(* IEC 61131-3 sources: 2026_Projet_YGO_ExcavatriceDragage/CODE_BACKUP/CODE_20260907_ChantierWeekEnd_v0.6.43/J_SUPERVISION/_TYPES/1_TREUILS_BENNE, 26 files *)

(* ---- E_WinchTraceBlockReason.st ---- *)
(* =======================================================================
   E_WinchTraceBlockReason - Cause de blocage priorisee treuil (trace terrain)
   -----------------------------------------------------------------------
   Role : Ordre de priorite de la cause de blocage d'un treuil M1/M2,
      calcule en PRG_04_Treuils_Benne (#8bis) et publie via Data.TraceM1/M2.
      L'ordre de l'enum EST l'ordre de priorite (valeur croissante = priorite
      decroissante) : la cause la plus grave gagne (PowerCutOff > ... > NONE).
   Producteur unique : PRG_04_Treuils_Benne (#8bis).
   Consommateur : FB_TroubleshootingView (recopie -> GVL_Troubleshooting.TraceM1/2).
   Lecture seule - aucune action de conduite n'en depend.
   Doc metier : DOC/AF/AF_Partie-14_Fonction_Troubleshooting_v1.4.md
   ======================================================================= *)
{attribute 'qualified_only'}
TYPE E_WinchTraceBlockReason :
(
    NONE                    := 0,   // Aucun blocage - au moins un sens effectivement permis
    POWER_CUTOFF            := 1,   // Coupure puissance amont (instSafetyWinch.PowerCutOff) - priorite max
    AXIS_DISABLED           := 2,   // Axe neutralise (Mode=DISABLE ou InhibitMx -> Enable FALSE)
    SAFESTOP                := 3,   // SafeStop effectif (rampe rapide demandee)
    SAFETY_FAULT            := 4,   // Defaut safety latched (FB_Safety_Winch.Fault.Error)
    SAFETY_PERMIT_MISSING   := 5,   // Aucun sens ne delivre de permit safety (limite / mou de cable / homing)
    PROCESS_PERMIT_MISSING  := 6,   // Permit process absent (benne / fond Kobold / limite legale / extraction)
    COUPLING_BLOCKED        := 7,   // Couplage synchro anti-telescopage (l'autre axe bloque)
    WINCH_FAULT             := 8,   // Defaut treuil latched (FB_Winch.Fault.Error)
    FINAL_INTERLOCK_BLOCKED := 9    // Barriere finale en defaut (frein / redemarrage)
);
END_TYPE

(* ---- ST_BucketCfg.st ---- *)
(* ═══════════════════════════════════════════════════════════════
   ST_BucketCfg — Configuration de la benne (M2)
   ═══════════════════════════════════════════════════════════════ *)
TYPE ST_BucketCfg :
STRUCT
    Config              : ST_fbBucket_Config; (* Offsets Open/Close/Coherence *)
    CfgTimeoutDuration  : TIME := T#30s;    (* ⏱️ Temps max pour l'ouverture/fermeture *)
    Initialized         : BOOL := FALSE;   (* 🚦 flag restauration boot *)
END_STRUCT
END_TYPE

(* ---- ST_BucketCmd.st ---- *)
(* ═══════════════════════════════════════════════════════════════
   🎮 ST_BucketCmd — Commandes IHM pour la benne (M2)
   ═══════════════════════════════════════════════════════════════ *)
TYPE ST_BucketCmd :
STRUCT
    BtnOpen             : BOOL; (* 🪣 Bouton commande ouverture *)
    BtnClose            : BOOL; (* 🪣 Bouton commande fermeture *)
    BtnReset            : BOOL; (* 🔑 Acquittement défaut benne *)
    BtnConfirmOpenPos   : BOOL; (* Référencement benne position ouverte (mise en service) — confirmation pure, aucun mouvement *)
    BtnConfirmClosePos  : BOOL; (* Référencement benne position fermée (mise en service) — confirmation pure, aucun mouvement *)
    // Mode pilotage unitaire M2 "sécurisé" -- actif
    // uniquement en SelJoystickWinch=2 (unitaire M2). Si TRUE : borne le déplacement entre les
    // positions ouvert/fermé configurées (OffsetOpenM/OffsetCloseM relatif à M1, mêmes bornes que
    // FB_Bucket) ET plafonne la vitesse au palier 1, sans passer par instBucket (pas de mémorisation
    // CloseReq/OpenReq, jogging libre borné). Défaut FALSE : pilotage unitaire M2 sans limite dédiée.
    TglManualBucketLimits : BOOL := TRUE; // Défaut TRUE -- pilotage unitaire M2 borné + palier 1 par défaut
    // Assistance "vidage à la trémie" (MAINT_N1/N2) : arme l'ouverture auto de la benne quand
    // M3 est stable à la Trémie. Indépendant du verrou descente treuil (WinchDescentAuth_M3).
    TglEnableDumpAtTremie : BOOL := FALSE;
END_STRUCT
END_TYPE

(* ---- ST_BucketHMI.st ---- *)
(* ═══════════════════════════════════════════════════════════════
   ⚙️ ST_BucketHMI — Données d'échange IHM pour la benne (M2)
   ───────────────────────────────────────────────────────────────
   📄 Structuration en Cmd / State / Cfg / Bypass , homogène avec ST_WinchHMI.
   ═══════════════════════════════════════════════════════════════ *)
TYPE ST_BucketHMI :
STRUCT
    Cmd    : ST_BucketCmd;
    State  : ST_BucketHMIState;
    Cfg    : ST_BucketCfg;
    Bypass : ST_BypassBucket;
END_STRUCT
END_TYPE

(* ---- ST_BypassBucket.st ---- *)
(* ═══════════════════════════════════════════════════════════════
   ST_BypassBucket — Bypass de la surveillance benne (M2)
   🔒 Doctrine : actionnable UNIQUEMENT en MAINT_N2, RETAIN, jamais masque
      les autres défauts du même bloc.
   ═══════════════════════════════════════════════════════════════ *)
TYPE ST_BypassBucket :
STRUCT
    (* 🛡️ 1. Hiérarchie & Restauration *)
    Global      : BOOL; (* 🌐 Bypass Global : ignore toute surveillance du mécanisme benne *)
    // Flag restauration boot dédié (défaut FALSE non ambigu, contrairement à une valeur métier)
    Initialized : BOOL := FALSE; (* 🚦 TRUE = bypass restauré depuis GVL_BypassRetain ce boot *)
END_STRUCT
END_TYPE

(* ---- ST_BypassWinch.st ---- *)
(* ═══════════════════════════════════════════════════════════════
   ST_BypassWinch — Bypass maintenance dédiés à UN treuil (M1 ou M2)
   ───────────────────────────────────────────────────────────────
   🎨 Regroupe les bypass "dégradé assumé" propres à un axe (codeur,
      contacteurs) — chaque treuil a son propre matériel, donc son
      propre struct (imbriqué M1Winch.Bypass / M2Winch.Bypass).
   🔒 Doctrine : actionnable UNIQUEMENT en MAINT_N2, RETAIN, jamais masque
      les autres défauts du même bloc (voir REGISTRE_ACTIONS_Bypass_v1.0 (archive)).
   ⚠️ Les bypass de capteurs COMMUNS (SlackCable, TopPositionSensor — capteur
      physique unique partagé M1/M2) sont dans ST_CommunHMI.Bypass, PAS ici.
   ═══════════════════════════════════════════════════════════════ *)
TYPE ST_BypassWinch :
STRUCT
    (* 📡 1. Communication & Systèmes auxiliaires *)
    OperatorComm      : BOOL; (* 📡 Bypass communication esclave CANopen Joystick / heartbeat IHM *)
    EncoderFault      : BOOL; (* 🔌 Bypass diagnostic esclave EtherCAT COD (codeur absolu) *)
    ContactorFeedback : BOOL; (* 🔌 Bypass feedbacks contacteurs de puissance et frein *)
    PhaseRotation     : BOOL; (* ⚡ Bypass défaut rotation de phases (commun machine) *)
    BrakeThermal      : BOOL; (* 🌡️ Bypass surchauffe thermique frein (commun machine) *)
    MotorThermal      : BOOL; (* : 🌡️ Bypass surchauffe thermique moteur CE treuil (M1_ThermalOk_DI/M2_ThermalOk_DI) *)

    (* 🚧 2. Limites physiques et Positionnement *)
    TopLimitSwitch    : BOOL; (* 🚧 Bypass fin de course physique haute (capteur, bit5) *)
    TopLimitSoftware  : BOOL; (* : Bypass fin de course logiciel haut (position calculée CablePosM >= TopLimitM, symétrique CableLimitSwitch) *)
    CableLimitSwitch  : BOOL; (* 🚧 Bypass limite basse physique (longueur de câble max) *)
    LimitLegal        : BOOL; (* : Bypass limite légale de profondeur (GVL_IHM.Commun.LimitLegalReached) *)

    (* ⚙️ 3. Sécurité Mécanique (Méca A-E) *)
    MecaA             : BOOL; (* 🔄 Bypass Méca A : mouvement non commandé à l'arrêt *)
    MecaB             : BOOL; (* 🛑 Bypass Méca B : absence confirmation arrêt (frein/contacteurs) *)
    MecaC             : BOOL; (* 🏋️ Bypass Méca C : glissement de charge (benne M1) *)
    MecaD             : BOOL; (* 🚧 Bypass Méca D : arrivée butée haute anormale *)
    MecaE             : BOOL; (* 🔄 Bypass Méca E : désynchronisation critique *)

    (* 🛡️ 4. Hiérarchie & Restauration *)
    Safety            : BOOL; (* 🛡️ Bypass groupé : tous les bits qui provoquent un PowerCutOff *)
    Process           : BOOL; (* ⚙️ Bypass groupé : tous les bits qui provoquent un SafeStop *)
    Global            : BOOL; (* 🌐 Bypass Global : ignore toutes les sécurités de cet axe *)
    // Flag restauration boot dédié (défaut FALSE non ambigu, contrairement à une valeur métier)
    Initialized       : BOOL := FALSE; (* 🚦 TRUE = bypass restauré depuis GVL_BypassRetain ce boot *)
END_STRUCT
END_TYPE

(* ---- ST_Chain_Winch_Control.st ---- *)
TYPE ST_Chain_Winch_Control :
STRUCT
    Idx401_MotionAllowed         : BOOL; // 1 = Prêt / Mouvement Autorisé | 0 = Bloqué
    Idx402_SpeedStepCalculated   : INT;  // Palier Vitesse Calculé (0, 1, 2, 3, 4)
    Idx403_SpeedRamp_Pct         : REAL; // [%] Consigne Vitesse après Rampe
    Idx404_BrakeReleaseAuthorized: BOOL; // 1 = Ordre Ouverture Frein | 0 = Ordre Serrage
    Idx405_FinalInterlockState   : E_WinchFinalInterlockState; // 🛡️ État frontière
    Idx406_FinalInterlockReason  : E_WinchFinalInterlockReason; // 🛡️ Cause mémorisée
    Idx407_FinalAuthorizedStep   : INT;  // 🪜 Palier réellement autorisé
    Idx408_BrakeCommandOpenConfirmed : BOOL; // 🔌 Contacteur/bobine, pas frein mécanique
    Idx409_BrakeTimeoutElapsed   : TIME; // ⏱️ Watchdog 500ms écoulé
    Idx410_RestartDelayElapsed   : TIME; // ⏱️ Verrou 900ms écoulé
    Idx411_StepDelayElapsed      : TIME; // ⏱️ Délai palier 1s250 écoulé
    Idx412_InTopSlowdownZone     : BOOL; // 🐢 Palier plafonné à 1, approche limite haute
    Idx413_InBottomSlowdownZone  : BOOL; // 🐢 Palier plafonné à 1, approche limite basse (câble ou légale)
    Idx414_BottomLimitActiveM    : REAL; // : Limite basse active (m) — câble physique OU légale, la plus restrictive
    (* 🔎 Diagnostic anti-redémarrage — "commande active mais rien ne tourne" *)
    Idx415_MotorRequest          : BOOL; // 1 = demande moteur active (palier>0 ET un seul sens) | 0 = pas de demande vue par la barrière
    Idx416_RestartRequired       : BOOL; // 1 = purge anti-redémarrage armée, AuthorizedStep force a 0 tant que non purgee
    Idx417_RestartInhibit        : BOOL; // 1 = verrou latché (frein non confirmé), exige Reset conscient — distinct de Idx416
    Idx418_NeutralRequestSeen    : BOOL; // 1 = passage au neutre observé pendant un RestartInhibit (réarmement en cours)
END_STRUCT
END_TYPE

(* ---- ST_Chain_Winch_Demandes.st ---- *)
TYPE ST_Chain_Winch_Demandes :
STRUCT
    Idx201_JoyRawPhysical_ANA    : INT;  // [pts] Bruts convertisseur (-2048 à +2048)
    Idx202_JoyScaledPhysical_Pct : REAL; // [%] Consigne Joystick (-100% à +100%)
    Idx203_HmiManualCmd_BtnAscent : BOOL; // 1 = Appui Bouton Ascending IHM | 0 = Relâché
    Idx204_HmiManualCmd_BtnDescent : BOOL; // 1 = Appui Bouton Descending IHM | 0 = Relâché
    Idx205_CycleAutoCmd_Pct      : REAL; // [%] Consigne auto envoyée par le Cycle
    Idx206_ModeActive            : E_Mode;// Mode courant (MANU_N1, AUTO_N1, MAINT_N2...)
    Idx207_BypassOperatorComm    : BOOL; // 0 = Comm Normale OK | 1 = Bypass Réseau Actif ⚠️
    Idx208_ArbitratedSpeed_Pct   : REAL; // [%] Consigne finale retenue après arbitrage
    Idx209_ArbitratedDirection   : INT;  // +1 = Ascending | 0 = Neutre | -1 = Descending
    Idx210_CoupledUserRequestDirection : INT; // +1 = Ascending | 0 = Neutre | -1 = Descending
    Idx211_CoupledUserRequestActive    : BOOL; // 1 = demande utilisateur couplée active
END_STRUCT
END_TYPE

(* ---- ST_Chain_Winch_Inputs.st ---- *)
TYPE ST_Chain_Winch_Inputs :
STRUCT
    Idx101_EncoderRawPos         : DINT; // [Valeur brutes pts] Codeur connecté
    Idx102_CablePos_M            : REAL; // [mètres] Position calculée du câble
    Idx103_ContactorsReleased_DI : BOOL; // 1 = OK (Tous contacteurs retombés à l'arrêt) | 0 = Contacteur collé
    Idx104_BrakeApplied          : BOOL; // TRUE = frein SERRÉ (NOT BrakeFeedback — IHM garde le sens serré)
    Idx105_ThermalOk_DI          : BOOL; // 1 = Température OK (Sain) | 0 = Surchauffe Moteur M1
END_STRUCT
END_TYPE

(* ---- ST_Chain_Winch_Outputs.st ---- *)
TYPE ST_Chain_Winch_Outputs :
STRUCT
    Idx501_CmdRelayAscent_DQ   : BOOL; // 1 = Relais Ascending ON | 0 = OFF
    Idx502_CmdRelayDescent_DQ  : BOOL; // 1 = Relais Descending ON | 0 = OFF
    Idx503_CmdSpeedContactor1_DQ : BOOL; // 1 = Contacteur Vitesse 1 ON | 0 = OFF
    Idx504_CmdSpeedContactor4_DQ : BOOL; // 1 = Contacteur Vitesse 4 ON (Plein Gaz) | 0 = OFF
    Idx505_CmdBrakeRelease_RQ    : BOOL; // 1 = Bobine Frein Alimentée (Ouvert) | 0 = Non Alimentée (Serré)
END_STRUCT
END_TYPE

(* ---- ST_Chain_Winch_Safety.st ---- *)
TYPE ST_Chain_Winch_Safety :
STRUCT
    Idx301_EmergencyChainClosed  : BOOL; // 1 = Boucle Urgence OK (Armé) | 0 = Arrêt d'Urgence Appuyé
    Idx302_SafeStopActive        : BOOL; // 0 = Sain (Autorisé) | 1 = Arrêt Rapide Métier Actif
    Idx303_PowerCutOffActive     : BOOL; // 0 = Puissance OK | 1 = Coupure Puissance Sécurité
    Idx304_TopSensorPhysical_DI  : BOOL; // 1 = Capteur Haut Libre (Sain) | 0 = Butée Haute Atteinte
    Idx305_TopSensorBypassActive : BOOL; // 0 = Capteur Actif | 1 = Capteur Haut Shunté IHM ⚠️
    Idx306_AscentPermitEffective  : BOOL; // 1 = Ascending Autorisée | 0 = ASCENDING BLOQUÉE
    Idx307_SlackCablePhysical_DI : BOOL; // 1 = Câble Tendu (Sain) | 0 = Mou de Câble Détecté
    Idx308_SlackCableBypassActive: BOOL; // 0 = Capteur Actif | 1 = Mou de Câble Shunté IHM ⚠️
    Idx309_DescendPermitEffective: BOOL; // 1 = Descending Autorisée | 0 = DESCENDING BLOQUÉE
    (* Défauts safety déchiffrés (bits ErrorId) — visibles individuellement à l'IHM *)
    Idx310_ErrorOperatorComm : BOOL; // bit0 Perte communication opérateur (joystick CAN / heartbeat IHM)
    Idx311_ErrorEncoder      : BOOL; // bit1 Perte codeur de ce treuil
    Idx312_ErrorPhaseRotation: BOOL; // bit4 Mauvaise rotation de phases
    Idx313_ErrorMecaA        : BOOL; // bit7 Mouvement non commandé / roue libre
    Idx314_ErrorMecaB        : BOOL; // bit8 Absence confirmation arrêt sans commande
    Idx315_ErrorMecaC        : BOOL; // bit9 Glissement M1 pendant cycle benne
    Idx316_ErrorMecaD        : BOOL; // bit11 Non-arrêt sur capteur haut
    Idx317_ErrorMecaE        : BOOL; // bit12/13 Écart synchro critique M1/M2
    Idx318_ErrorBrakeThermal : BOOL; // bit10 Surchauffe thermique frein commun
    Idx319_ErrorOppositeDir  : BOOL; // bit14 Sens réel opposé au sens commandé
    Idx320_ErrorNoMovement   : BOOL; // bit15 Absence de mouvement malgré commande
    (* ⛔ Bloc "Pourquoi la montée ne s'arrête pas à la limite haute ?" — diagnostic ordonné
       (lecture maintenance) : config + position → butée atteinte → bypass actifs. *)
    Idx321_CfgTopLimitM               : REAL;  // 📐 Limite haute effective active (m) = CfgCableLimitAscent_M
    Idx322_CablePosM                  : REAL;  // 📐 Position câble courante (m)
    Idx323_TopLimitReached            : BOOL;  // 1 = position >= limite haute (hors homing) | 0 = en dessous
    Idx324_AscentBlockedByTopLimit    : BOOL;  // 1 = montée réellement coupée par la butée logicielle (AscentPermit=0) | 0 = limitée non bloquante (bypass ?)
    Idx325_BypassTopLimitSoftware     : BOOL;  // ⚠️ 1 = butée logicielle shunétee IHM (individuel)
    Idx326_BypassTopLimitSoftCommun   : BOOL;  // ⚠️ 1 = butée logicielle shunétee (commun)
    Idx327_BypassTopLimitSwitch       : BOOL;  // ⚠️ 1 = capteur fin de course haut shuné IHM (individuel)
    Idx328_BypassTopLimitSwitchCommun : BOOL;  // ⚠️ 1 = capteur fin de course haut shuné (commun)
    Idx329_BypassGlobal               : BOOL;  // ⚠️ 1 = bypass global treuil (individuel)
    Idx330_BypassGlobalCommun         : BOOL;  // ⚠️ 1 = bypass global (commun)
END_STRUCT
END_TYPE

(* ---- ST_ChainBucket.st ---- *)
TYPE ST_ChainBucket :
STRUCT
    Idx101_BucketIsOpen          : BOOL; // 1 = Benne Mécaniquement Ouvert | 0 = Non Confirmé
    Idx102_BucketIsClosed        : BOOL; // 1 = Benne Mécaniquement Fermé | 0 = Non Confirmé
    Idx103_OffsetPos_M           : REAL; // [mètres] Écart d'Ouverture Câble M1/M2
    Idx104_AutoSeqActive         : BOOL; // : 1 = Séquencement auto (ouverture/fermeture armée par mouvement couplé) en cours
    Idx105_StateIncoherent       : BOOL; // : 1 = État ouvert/fermé INCONNU (ni IsOpen ni IsClosed fiable) -- cause fréquente de blocage
    Idx106_FBState               : E_State; // : État machine FB_Bucket (READY/BUSY/DONE/DISABLED)
    Idx107_LastPosM2Open_M       : REAL; // : Dernière position M2 mémorisée "ouvert"
    Idx108_LastPosM2Close_M      : REAL; // : Dernière position M2 mémorisée "fermé"
    Idx109_BucketTooOpen         : BOOL; // ⚠️ Dépassement ouverture : Delta < OffsetOpen - Tolerance (Enrouler M2)
    Idx110_BucketTooClosed       : BOOL; // ⚠️ Dépassement fermeture : Delta > OffsetClose + Tolerance (Dérouler M2)
    Idx111_BucketIsIntermediate  : BOOL; // ↔️ Position intermédiaire (entrebâillée entre ouvert et fermé)
    Idx112_DeltaPosition_M       : REAL; // 📏 Écart réel signé M2 - M1 (mètres) en direct

    Idx113_MachineHomed : BOOL; // Reference M1/M2/benne qualifiee
    Idx114_MachineHomingStep         : INT;  // Etape guidee reference machine
    Idx115_MachineHomingFailed       : BOOL; // Transaction reference abandonnee
    Idx116_M1ReferenceMissing    : BOOL; // M1 non reference ou mesure douteuse
    Idx117_M2ReferenceMissing    : BOOL; // M2 non reference ou mesure douteuse
    Idx118_BucketOffsetUnknown   : BOOL; // Offset benne non confirme
    Idx119_ReferenceTransaction  : BOOL; // Homing conjoint en cours
    Idx120_MachineHomingLossSafeStop : BOOL; // Perte reference pendant mouvement

    Idx201_HmiCmd_BtnOpen        : BOOL; // 1 = Demande Ouverture IHM | 0 = Relâché
    Idx202_HmiCmd_BtnClose       : BOOL; // 1 = Demande Fermeture IHM | 0 = Relâché
    Idx203_CycleCmd_Open         : BOOL; // 1 = Demande Ouverture par le Cycle Auto
    Idx204_CoupledDiveOpenArmed   : BOOL; // : 1 = Ouverture auto armée (descente couplée demandée, benne pas ouverte)
    Idx205_CoupledAscentCloseArmed: BOOL; // : 1 = Fermeture auto armée (montée couplée demandée, benne pas fermée)
    Idx206_CloseReqActive        : BOOL; // : 1 = Fermeture mémorisée/en cours (instBucket.CloseReq -- reste à 1 si recul partiel non terminé)
    Idx207_OpenReqActive         : BOOL; // : 1 = Ouverture mémorisée/en cours (instBucket.OpenReq -- idem)
    Idx208_MotionBlockedByBucket : BOOL; // : 1 = Mouvement couplé BLOQUÉ (auto-séquencement armé mais benne pas Busy -- vérifier Idx306_ErrorIdRaw)

    Idx301_EmergencyChainClosed  : BOOL; // 1 = Boucle Urgence OK | 0 = AU Appuyé
    Idx302_BucketFaultActive     : BOOL; // 0 = Sain | 1 = Défaut Mouvement Benne
    Idx303_KoboldAutoStopEnabled       : BOOL; // 1 = Toggle IHM arrêt auto descente actif
    Idx304_KoboldImmersionConfirmed    : BOOL; // : 1 = Immersion confirmée (front Kobold dans la fenêtre)
    Idx305_KoboldBottomTouchLatched    : BOOL; // : 1 = Fond détecté, descente bloquée (ProcessPermitM1/M2_Descend)
    Idx306_ErrorIdRaw             : WORD; // : bitfield brut FB_Bucket (bit0 configuration, bit1 écart M2/M1, bit2 timeout, bit3 glissement M1, bit4 codeurs non référencés)
    Idx307_EffectivePermit_Open    : BOOL; // 1 = ouverture benne physiquement autorisée
    Idx308_EffectivePermit_Close   : BOOL; // 1 = fermeture benne physiquement autorisée

    Idx401_BucketBusy            : BOOL; // 1 = Mouvement Mâchoires en cours | 0 = Repos
    Idx402_BucketDone            : BOOL; // 1 = Position Cible Atteinte | 0 = En cours
    Idx403_ExtractionControlActive : BOOL; // : 1 = Phase vitesse contrôlée montée en cours

    Idx501_M2_CmdRev_DQ          : BOOL; // 1 = Relais Action Benne M2 ON
END_STRUCT
END_TYPE

(* ---- ST_ChainWinch.st ---- *)
TYPE ST_ChainWinch :
STRUCT
    Inputs_100    : ST_Chain_Winch_Inputs;
    Demandes_200  : ST_Chain_Winch_Demandes;
    Safety_300    : ST_Chain_Winch_Safety;
    Control_400   : ST_Chain_Winch_Control;
    Outputs_500   : ST_Chain_Winch_Outputs;
END_STRUCT
END_TYPE

(* ---- ST_ChainWinchSync.st ---- *)
TYPE ST_ChainWinchSync :
STRUCT
    Idx101_M1_CablePos_M         : REAL; // [mètres] Position Câble M1 Retenue
    Idx102_M2_CablePos_M         : REAL; // [mètres] Position Câble M2 Benne
    Idx103_SyncDelta_M           : REAL; // [mètres] Écart Relatif M1 - M2

    Idx201_JoyYRaw_Pct           : REAL; // [%] Consigne Joystick Axe Y (-100% à +100%)
    Idx202_SyncEnabled_IHM       : BOOL; // 1 = Couplage Synchro Actif (Nominal) | 0 = Découplé ⚠️
    Idx203_ArbitratedSpeed_Pct   : REAL; // [%] Consigne Vitesse Synchro Arbitrée

    Idx301_EmergencyChainClosed  : BOOL; // 1 = Boucle Urgence OK | 0 = Arrêt Urgence
    Idx302_SyncFaultActive       : BOOL; // 0 = Synchro OK | 1 = Écart Synchro Bloquant
    Idx303_M1_AscentPermit       : BOOL; // 1 = Ascending M1 Autorisée | 0 = Bloquée (Fdc/Safety)
    Idx304_M2_AscentPermit       : BOOL; // 1 = Ascending M2 Autorisée | 0 = Bloquée (Fdc/Safety)

    Idx401_SyncMotionAllowed     : BOOL; // 1 = Mouvement Synchro Autorisé | 0 = Bloqué
    Idx402_M1_SetpointSpeed_Pct  : REAL; // [%] Consigne Vitesse Calculée M1
    Idx403_M2_SetpointSpeed_Pct  : REAL; // [%] Consigne Vitesse Calculée M2

    Idx501_M1_CmdRelayFwd_DQ     : BOOL; // 1 = Ascending M1 ON | 0 = OFF
    Idx502_M2_CmdRelayFwd_DQ     : BOOL; // 1 = Ascending M2 ON | 0 = OFF
END_STRUCT
END_TYPE

(* ---- ST_HwWinch.st ---- *)
(* ═══════════════════════════════════════════════════════════════
   🏗️ ST_HwWinch — Image matérielle brute des entrées Treuils M1 / M2
   ───────────────────────────────────────────────────────────────
   🎨 Regroupe les signaux physiques d'entrée bruts des treuils M1 et M2.
   ═══════════════════════════════════════════════════════════════ *)
TYPE ST_HwWinch :
STRUCT
    M1_ContactorsReleased_DI : BOOL; (* Retours contacteurs M1 retombés *)
    M1_ThermalOk_DI          : BOOL; (* Thermique moteur M1 OK *)
    M1_BrakeIsOpen_DI        : BOOL; (* Retour frein M1 (1 = ouvert) *)

    M2_ContactorsReleased_DI : BOOL; (* Retours contacteurs M2 retombés *)
    M2_ThermalOk_DI          : BOOL; (* Thermique moteur M2 OK *)
    M2_BrakeIsOpen_DI        : BOOL; (* Retour frein M2 (1 = ouvert) *)

    M1M2_TopPositionFree_DI  : BOOL; (* Capteur position haute commun M1/M2 libre *)
    M2_TensionedCable_DI     : BOOL; (* Capteur mou de câble M2 (câble tendu) *)

    COD1_PosValue            : UDINT;        (* Valeur brute position codeur COD1 (M1) *)
    COD1_SpdValue            : DINT;         (* Valeur brute vitesse codeur COD1 (0x6031:01 en 0.1 RPM) *)
    COD1_Alarms              : UINT;         (* Alarmes brutes COD1 *)
    COD1_Warnings            : UINT;         (* Avertissements bruts COD1 *)
    COD1_DeviceState         : DEVICE_STATE; (* État device COD1 (GetDeviceState) *)

    COD2_PosValue            : UDINT;        (* Valeur brute position codeur COD2 (M2) *)
    COD2_SpdValue            : DINT;         (* Valeur brute vitesse codeur COD2 (0x6031:01 en 0.1 RPM) *)
    COD2_Alarms              : UINT;         (* Alarmes brutes COD2 *)
    COD2_Warnings            : UINT;         (* Avertissements bruts COD2 *)
    COD2_DeviceState         : DEVICE_STATE; (* État device COD2 (GetDeviceState) *)
END_STRUCT
END_TYPE

(* ---- ST_OutputsInterPrg.st ---- *)
(* ═══════════════════════════════════════════════════════════════
   📤 ST_OutputsInterPrg — Bus d'échange inter-PRG produit par PRG_06_Outputs
   ───────────────────────────────────────────────────────────────
   🎯 Rôle : Encapsuler les ordres actionneurs finaux (M1/M2/M3, AU) produits
      par PRG_06_Outputs et rebouclés par FB_SimBench (instancié dans
      PRG_02_Acquisition) pour le banc de simulation intégré.
   📤 Producteur unique : PRG_06_Outputs (VAR_OUTPUT Data : ST_OutputsInterPrg).
   📄 Doc : DOC/AF/AF_Partie-06_Acquisition_Qualification_IO_v2.4.md §5
   🔌 Architecture : Bus de données typé — encapsulation des échanges inter-PRG.
   ═══════════════════════════════════════════════════════════════ *)

TYPE ST_OutputsInterPrg :
STRUCT
    // === 🪝 Ordres actionneurs finaux treuil M1 ===
    M1RelayFwd            : BOOL; // 🛗 Ordre contacteur montee treuil M1
    M1RelayRev            : BOOL; // 🛗 Ordre contacteur descente treuil M1
    M1SpeedContactor1     : BOOL; // 🔌 Ordre contacteur palier 1 treuil M1
    M1SpeedContactor2     : BOOL; // 🔌 Ordre contacteur palier 2 treuil M1
    M1SpeedContactor3     : BOOL; // 🔌 Ordre contacteur palier 3 treuil M1
    M1SpeedContactor4     : BOOL; // 🔌 Ordre contacteur palier 4 treuil M1
    M1BrakeCmd            : BOOL; // 🔓 Ordre desserrage frein M1 (1=Desserrer)

    // === 🪝 Ordres actionneurs finaux treuil M2 ===
    M2RelayFwd            : BOOL; // 🛗 Ordre contacteur montee/fermeture treuil M2
    M2RelayRev            : BOOL; // 🛗 Ordre contacteur descente/ouverture treuil M2
    M2SpeedContactor1     : BOOL; // 🔌 Ordre contacteur palier 1 treuil M2
    M2SpeedContactor2     : BOOL; // 🔌 Ordre contacteur palier 2 treuil M2
    M2SpeedContactor3     : BOOL; // 🔌 Ordre contacteur palier 3 treuil M2
    M2SpeedContactor4     : BOOL; // 🔌 Ordre contacteur palier 4 treuil M2
    M2BrakeCmd            : BOOL; // 🔓 Ordre desserrage frein M2 (1=Desserrer)

    // === 🔀 Concordance contacteurs M1/M2 (instance FB_SyncContactor sur vecteurs finaux) ===
    ContactorMismatch          : BOOL;                  // Niveau 1 confirmé (debounce 500 ms) → SafeStop des 2 treuils (PRG_04, scan N-1)
    ContactorMismatchEscalated : BOOL;                  // Niveau 2 persistant → escalade PowerCutOff via latch MecaE (PRG_04)
    SyncContactorDiag          : ST_SyncContactorDiag;  // Détail : quel contacteur diverge + niveau atteint (IHM / troubleshooting)

    // === ↔️ Ordre actionneur final translation M3 ===
    TranslationBrakeCmd   : BOOL; // 🔓 Demande frein M3 arbitree

    // === 🚨 Chaîne réarmement puissance AU ===
    PowerKeepAliveACmd    : BOOL; // 🔒 Maintien puissance voie A (1=Maintenu)
    PowerKeepAliveBCmd    : BOOL; // 🔒 Maintien puissance voie B (1=Maintenu)
    EmergencyArmingCmd    : BOOL; // 🎯 Impulsion rearmement puissance AU
    TestCutActive         : BOOL; // 🧪 Test de redondance AU en cours (canal A ou B coupe) — consommé par FB_SimBench
    PowerCutOffRequest    : BOOL; // 🛑 Requête coupure métier (arrêt d'urgence) — consommé par FB_SimBench
END_STRUCT
END_TYPE

(* ---- ST_SafetyWinch.st ---- *)
(* ═══════════════════════════════════════════════════════════════
   🛡️ ST_SafetyWinch — Diagnostics de sécurité pour un treuil
   ───────────────────────────────────────────────────────────────
   🎨 Destiné à l'affichage des défauts de sécurité d'un treuil.
   ═══════════════════════════════════════════════════════════════ *)
TYPE ST_SafetyWinch :
STRUCT
    Error             : BOOL;    (* 🛡️ Bloc sécurité (Safety) en défaut *)
    ErrorId           : WORD;    (* ❌ Code bitfield du défaut de sécurité (vue LIVE) *)
    LatchedId         : WORD;    (* 🕘 Vue LATCHÉE : ErrorId figé au défaut, effacé au Reset (marqueur [HISTO]) *)
    SafeStop          : BOOL;    (* 🟧 Arrêt rapide activé par la sécurité *)
    DescendPermit     : BOOL;    (* 🟢 Descending autorisée (TRUE = OK | FALSE = mou de câble / limite basse) *)
    AscentPermit      : BOOL;    (* 🟢 Ascending autorisée (TRUE = OK | FALSE = fin de course haut) *)
    SlackCable        : BOOL;    (* ⚠️ Mou de câble physiquement détecté *)
    ThermalFault      : BOOL;    (* 🔥 Surchauffe thermique moteur *)
    EncoderFault      : BOOL;    (* 🔌 Perte de liaison ou incohérence codeur *)
    BypassActive      : BOOL;    (* Bypass codeur effectivement accepté, uniquement MAINT_N2 *)
    CableLimitDescent : BOOL;    (* ⚠️ Longueur max de câble atteinte (limite basse physique) *)
    CableLimitAscent  : BOOL;    (* ⚠️ Limite haute d'exploitation normale atteinte *)
    MecaADrift_M      : REAL;    (* 📐 Dérive mesurée Méca A (m) *)
    MecaCDrift_M      : REAL;    (* 📐 Dérive mesurée Méca C (m) *)
    MecaBElapsedTime  : TIME;    (* ⏳ Temps écoulé confirmation contacteurs/frein *)
    PowerCutOff       : BOOL;    (* 🧨 Coupure puissance amont activée *)
    BlockedBySafety   : BOOL;    (* 🚫 Synthèse globale : actionneur bloqué par la sécurité (PowerCutOff OU SafeStop/Error) *)
    PowerCutOffSafety : BOOL;    (* 🧨 Synthèse sécurités critiques entraînant une coupure puissance *)
    SafeStopSafety    : BOOL;    (* 🛡️ Synthèse défauts entraînant un SafeStop / Rampe rapide *)
    (* 🔍 Décomposition individuelle des défauts de sécurité (bits ErrorId) *)
    ErrorOperatorComm : BOOL;    (* 🎮 Perte communication opérateur : joystick CAN ou heartbeat IHM (bit0) *)
    ErrorEncoder      : BOOL;    (* 🔌 Perte de liaison ou incohérence codeur (bit1) *)
    ErrorPhaseRotation: BOOL;    (* ⚡ Mauvaise rotation de phases électriques (bit4) *)
    ErrorBrakeThermal : BOOL;    (* 🌡️ Surchauffe thermique frein commun M1/M2/M3 (bit10) *)
    ErrorMecaA        : BOOL;    (* 🔄 Mouvement non commandé / roue libre (Méca A - bit7) *)
    ErrorMecaB        : BOOL;    (* 🛑 Absence confirmation arrêt sans commande (Méca B - bit8) *)
    ErrorMecaC        : BOOL;    (* 🏋️ Glissement M1 pendant cycle benne (Méca C - bit9) *)
    ErrorMecaD        : BOOL;    (* 🚧 Non-arrêt sur capteur haut (Méca D - bit11) *)
    ErrorMecaE        : BOOL;    (* 🔄 Écart de synchronisation critique M1/M2 (Méca E - bit12/13) *)
    ErrorOppositeDir  : BOOL;    (* 🧭 Sens réel opposé au sens commandé (bit14) *)
    ErrorNoMovement   : BOOL;    (* ⏱️ Absence de mouvement malgré commande (bit15) *)
    ErrorOverspeed    : BOOL;    (* ⚡ Survitesse treuil mesurée au-delà du palier 5 (latchée, acquittée au Reset) *)
END_STRUCT
END_TYPE

(* ---- ST_TraceWinch.st ---- *)
(* =======================================================================
   ST_TraceWinch - Trace de blocage terrain d'un treuil M1/M2
   -----------------------------------------------------------------------
   Role : Publier au technicien une vue consolidee "pourquoi l'axe ne bouge
   pas" : permis effectifs par sens, source du SafeStop/coupure, cause de
   blocage priorisee et horodatee.
   Producteur unique : PRG_04_Treuils_Benne (#8bis) - 1 instance par axe
       (TraceM1 / TraceM2 au sein de ST_WinchInterPrg).
   Consommateur : FB_TroubleshootingView (pure recopie -> GVL_Troubleshooting).
   Lecture seule - aucun calcul de commande n'en depend.
   BlockReasonTimestamp : ms depuis demarrage PLC (TIME()), latched au dernier
       changement de BlockReason (1 scan, memoire).
   Doc metier : DOC/AF/AF_Partie-14_Fonction_Troubleshooting_v1.4.md
   ======================================================================= *)
TYPE ST_TraceWinch :
STRUCT
    // Permis effectifs par sens (reflet exact des permis appliques au mouvement)
    DescendPermitEffective  : BOOL;   // Descente effectivement permise (EffectivePermit*_Descend)
    AscentPermitEffective   : BOOL;   // Montee effectivement permise (EffectivePermit*_Ascent)
    AscentPermitApplied      : BOOL;   // Permis effectivement transmis a la barriere finale
    DescendPermitApplied     : BOOL;   // Permis effectivement transmis a la barriere finale
    FinalPermitBlocked       : BOOL;   // Demande presente mais refusee par le permis final

    // Source de SafeStop / coupure - pour distinguer l'origine du blocage
    SafeStopActive          : BOOL;   // SafeStop effectif applique (SafeStop*_Active)
    SafeStopSourceSafety    : BOOL;   // SafeStop issu de FB_Safety_Winch (defaut safety)
    SafeStopSourceInput     : BOOL;   // SafeStop issu du module d'entree / homing / slip benne
    SafeStopSourceSync      : BOOL;   // SafeStop issu de la synchro M1/M2 (couplage anti-telescopage)
    PowerCutOffActive       : BOOL;   // Coupure puissance amont active (instSafetyWinch.PowerCutOff)
    Inhibited               : BOOL;   // Axe neutralise (Mode=DISABLE ou InhibitMx)

    // Barriere finale (fin de course mecanique / frein / redemarrage)
    FinalInterlockError     : BOOL;   // Defaut barriere finale (frein / redemarrage)
    FinalInterlockReason    : E_WinchFinalInterlockReason; // Cause barriere finale memorisee

    // Cause de blocage priorisee + horodatage
    BlockReason             : E_WinchTraceBlockReason; // Cause de blocage prioritaire
    BlockReasonTimestamp    : UDINT;  // ms depuis demarrage PLC (TIME()) - dernier changement de BlockReason
    StepNumber              : INT;    // Palier de vitesse actif (WinchState.StepNumber)
END_STRUCT
END_TYPE

(* ---- ST_WinchBenneHMI.st ---- *)
(* ═══════════════════════════════════════════════════════════════
   ⚙️ ST_WinchBenneHMI — Données d'échange IHM pour le treuil Benne (M2 uniquement)
   ───────────────────────────────────────────────────────────────
   🎨 Composition dupliquée de ST_WinchHMI (Cmd/State/Cfg/Safety/Bypass) + Bucket.
   📄 IEC 61131-3 n'offre pas d'héritage de struct : cette duplication de la liste
      de champs est assumée pour garder M1TreuilRetenue (ST_WinchHMI, sans Bucket)
      strictement distinct de M2TreuilBenne (ce type, avec Bucket) — décision
      DOC/CHECKLISTS/TASK_CONTEXT/TASK_CONTEXT_LOT_TROUBLESHOOTING_VIEW_ET_WINCHHMI.yaml AC5.
   ═══════════════════════════════════════════════════════════════ *)
TYPE ST_WinchBenneHMI :
STRUCT
    (* 🎮 Commandes opérateur *)
    Cmd                     : ST_WinchCmd;

    (* 🚦 États, retours et mesures *)
    State                   : ST_WinchState;

    (* Configurations et limites *)
    Cfg                     : ST_WinchCfg;

    (* 🛡️ Sécurité (FB_Safety_Winch) *)
    Safety                  : ST_SafetyWinch;

    (* Bypass maintenance *)
    Bypass                  : ST_BypassWinch;

    (* 🪣 Benne — pertinent uniquement pour M2 (M2TreuilBenne.Bucket) *)
    Bucket                  : ST_BucketHMI;
END_STRUCT
END_TYPE

(* ---- ST_WinchCfg.st ---- *)
(* ═══════════════════════════════════════════════════════════════
   ST_WinchCfg — Configurations et paramètres réglables pour un Treuil M1/M2
   ───────────────────────────────────────────────────────────────
   🎨 Destiné au paramétrage et calibration depuis l'IHM (RETAIN).
   ═══════════════════════════════════════════════════════════════ *)
TYPE ST_WinchCfg :
STRUCT
    CfgTopSensorPos_M       : REAL := 8.5;      (* 📐 Position cible du capteur haut (m) *)
    CfgHomingTarget_M       : REAL := 0.0;      (* Cible libre Homing unitaire MAINT_N2 [-99..+99 m] *)
    CfgRampAccelRate        : REAL := 50.0;     (* 📈 Rampe d'accélération (%/s) *)
    CfgRampDecelNormalRate  : REAL := 150.0;    (* 📉 Rampe de décélération normale (%/s) *)
    CfgRampDecelFastRate    : REAL := 400.0;    (* ⚡ Rampe de décélération rapide / SafeStop (%/s) *)
    CfgCableLimitDescent_M  : REAL := -50.0;    (* 📐 Limite basse physique de descente (m, négatif) *)

    (* 🚦 Flag restauration boot — défaut FALSE non ambigu *)
    Initialized              : BOOL := FALSE;    (* 🚦 TRUE = config restaurée depuis GVL_PERSISTENT ce boot *)
END_STRUCT
END_TYPE

(* ---- ST_WinchCmd.st ---- *)
(* ═══════════════════════════════════════════════════════════════
   🎮 ST_WinchCmd — Commandes IHM pour un Treuil M1/M2
   ───────────────────────────────────────────────────────────────
   🎨 Destiné au pilotage manuel et maintenance du treuil depuis l'IHM.
   ═══════════════════════════════════════════════════════════════ *)
TYPE ST_WinchCmd :
STRUCT
    BtnAscent               : BOOL;             (* ⬆️ Mouvement montee maintenu (mode boutons IHM, MAINT_N1 accessible) *)
    BtnDescent             : BOOL;             (* ⬇️ Mouvement descente maintenu (mode boutons IHM, MAINT_N1 accessible) *)
    BtnReset            : BOOL;             (* 🔑 Demande reset exposée par treuil ; agrégée dans le reset domaine partagé *)
    BtnHome             : BOOL;             (* 🎯 Homing nominal si Couplé, unitaire si M1/M2 sélectionné en MAINT_N2 *)
    BtnConfirmCoherence : BOOL;             (* 🔓 Confirmation de cohérence au démarrage *)
    BtnInhibit          : BOOL;             (* Bouton IHM inhibition treuil — mise en service,
                                                    UNIQUEMENT actif si MAINT_N2 (voir FB_Modes.InhibitM1/M2) *)
    BtnHomingAtZero     : BOOL;             (* Force le homing à 0 m (points codeur centre),
                                                    sans devoir modifier CfgTopSensorPos_M *)
    BtnOverrideTopSoftware : BOOL;          (* Autorisation MAINTENUE de dépasser le FDC
                                                    haut LOGICIEL (7,5 m) jusqu'au capteur physique
                                                    (CfgTopSensorPos_M ≈ 8,5 m). Bouton, pas toggle :
                                                    relâché ➔ retour immédiat à 7,5 m. Sans effet hors
                                                    MAINT_N1 (N2 utilise le bypass latché
                                                    Bypass.TopLimitSoftware). N'ouvre JAMAIS le FDC
                                                    capteur physique. *)
    BtnLearnSpeed : BOOL;                   (* 💾 Bit IHM lancer l'apprentissage passif des vitesses
                                                    réelles par palier (FB_WinchSpeedLearning).
                                                    Collecteur STRICTEMENT PASSIF : aucune commande moteur.
                                                    Maintenu pendant la collecte ; la table RETAIN
                                                    _WinchSpeedLearnTable est remplie par palier/sens/
                                                    charge/vide. *)
END_STRUCT
END_TYPE

(* ---- ST_WinchFinalInterlockRequest.st ---- *)
(* ═══════════════════════════════════════════════════════════════
   🪝 ST_WinchFinalInterlockRequest — Demande brute vers frontière Q M1/M2
   ───────────────────────────────────────────────────────────────
   📤 Producteur unique : PRG_04_Treuils_Benne (VAR_OUTPUT).
   📥 Consommateur unique : PRG_06_Outputs, avant FB_WinchOutputInterlock.
   🔒 Ne contient jamais une sortie Q autorisée : les C1..C4 restent les
      demandes exactes de FB_Winch / ST_SpeedStepTable.
   ═══════════════════════════════════════════════════════════════ *)

TYPE ST_WinchFinalInterlockRequest :
STRUCT
    Enable                       : BOOL;
    Reset                        : BOOL;
    PowerContactorEngaged              : BOOL;
    SafeStop                     : BOOL;
    BrakeFeedback                 : BOOL; // (retrait FB_Brake) : retour PHYSIQUE brut du
                                          // contacteur/bobine frein (TRUE = ouvert/relâché) — remplace
                                          // BrakeReleaseRequest/BrakeCommandOpenConfirmed ; la barrière
                                          // finale calcule elle-même BrakeCmd := RelayFwd OR RelayRev.
    FwdRevSpeedFeedbackOff       : BOOL; // TRUE = relais sens + C1..C4 tous retombés
    RequestedRelayFwd            : BOOL;
    RequestedRelayRev            : BOOL;
    RequestedContactor1          : BOOL;
    RequestedContactor2          : BOOL;
    RequestedContactor3          : BOOL;
    RequestedContactor4          : BOOL;
    RequestedStep                : INT;
    // Permis effectifs deja appliques par FB_Winch et reutilises par la barriere finale.
    AscentPermit                 : BOOL;
    DescendPermit                : BOOL;
    PowerCutOff                  : BOOL; // : demande coupure puissance (FB_Safety_Winch), agrégée par PRG_06 (M5, A-04)
END_STRUCT
END_TYPE

(* ---- ST_WinchHMI.st ---- *)
(* ═══════════════════════════════════════════════════════════════
   ⚙️ ST_WinchHMI — Données d'échange IHM pour un treuil (M1: moteur de retenue / M2: moteur Benne)
   ───────────────────────────────────────────────────────────────
   🎨 Destiné à l'affichage des bargraphes, LEDs, mesures et réglages.
   📄 Structuration en Cmd / State / Cfg / Safety / Bypass
   ═══════════════════════════════════════════════════════════════ *)
TYPE ST_WinchHMI :
STRUCT
    (* 🎮 Commandes opérateur *)
    Cmd                     : ST_WinchCmd;

    (* 🚦 États, retours et mesures *)
    State                   : ST_WinchState;

    (* Configurations et limites *)
    Cfg                     : ST_WinchCfg;

    (* 🛡️ Sécurité (FB_Safety_Winch) *)
    Safety                  : ST_SafetyWinch;

    (* Bypass maintenance *)
    Bypass                  : ST_BypassWinch;
END_STRUCT
END_TYPE

(* ---- ST_WinchInterPrg.st ---- *)
(* ═══════════════════════════════════════════════════════════════
   🪝 ST_WinchInterPrg — Bus d'échange inter-PRG produit par PRG_04_Treuils_Benne
   ───────────────────────────────────────────────────────────────
   🎯 Rôle : Encapsuler les demandes finales M1/M2, les états publics
      WinchM1/M2State, les sécurités WinchM1/M2Safety, l'état synchro et
      l'état benne publiés par PRG_04_Treuils_Benne vers les consommateurs
      (PRG_02/03/06/07).
   📤 Producteur unique : PRG_04_Treuils_Benne (VAR_OUTPUT Data : ST_WinchInterPrg).
   📄 Doc : DOC/AF/AF_Partie-10_Fonction_Winch_v2.1.md
   🔌 Architecture : Bus de données typé — encapsulation des échanges inter-PRG.
   ═══════════════════════════════════════════════════════════════ *)

TYPE ST_WinchInterPrg :
STRUCT
    // === ⚡ Demandes finales M1/M2 (interlocks & consigne vitesse arbitrée) ===
    WinchM1FinalInterlockRequest : ST_WinchFinalInterlockRequest; // 🪝 Demande finale et interlocks treuil M1
    WinchM2FinalInterlockRequest : ST_WinchFinalInterlockRequest; // 🪝 Demande finale et interlocks treuil M2
    M1LogicRequestSpeedCmd_Pct   : REAL; // 📈 Consigne vitesse M1 arbitree (%) — consommee par FB_SimBench (PRG_02)
    M2LogicRequestSpeedCmd_Pct   : REAL; // 📈 Consigne vitesse M2 arbitree (%) — consommee par FB_SimBench (PRG_02)
    KoboldContactorCmdArbitrated : BOOL; // 🪝 Ordre contacteur capteur fond Kobold (consommé PRG_06)

    // === 📊 États publics des treuils ===
    WinchM1State                 : ST_WinchState; // 🚦 Etat public treuil Retenue M1
    WinchM2State                 : ST_WinchState; // 🚦 Etat public treuil Benne M2

    // === 🛡️ Sécurités des treuils ===
    WinchM1Safety                : ST_SafetyWinch; // 🛡️ Diagnostic et securites treuil M1
    WinchM2Safety                : ST_SafetyWinch; // 🛡️ Diagnostic et securites treuil M2

    // === 🔄 État synchronisation ===
    SyncState                    : ST_SyncState; // 🔄 Etat synchronisation treuils M1/M2
    WinchSyncError               : BOOL;         // 🚨 Defaut de desynchronisme treuils M1/M2
    WinchSyncSignedDeltaPosM     : REAL;         // 📏 Ecart signe M2 - M1 (m)

    // === 🏗️ État benne ===
    BucketState                  : ST_BucketHMIState; // 🏗️ Etat de fonctionnement benne
    Benne_IsRoughlyClosed        : BOOL;               // 🏗️ Benne consideree fermee (tolerance matiere)
    BucketBusy                   : BOOL;               // ⚙️ Mouvement d'ouverture/fermeture benne en cours
    BucketDone                   : BOOL;               // ✅ Mouvement benne termine avec succes
    BucketError                  : BOOL;               // ❌ Defaut sur sous-systeme benne
    EffectivePermitBucket_Open   : BOOL;               // 🟢 Permis effectif ouverture benne
    EffectivePermitBucket_Close  : BOOL;               // 🟢 Permis effectif fermeture benne

    // === 🛡️ Permission d'armement homme-mort (Option B — combiné interlock benne) ===
    ArmingPermit                 : BOOL;               // 🛡️ Permission d'armement homme-mort (consommée PRG_02 → FB_Joystick). TRUE = armement autorisé (NC-100)
    ProcessPermitM1_Ascent       : BOOL;
    ProcessPermitM1_Descend      : BOOL;
    ProcessPermitM2_Ascent       : BOOL;
    ProcessPermitM2_Descend      : BOOL;
    DescendPermitDiveBucketOpen  : BOOL;
    ExtractionAssistActive       : BOOL;
    ExtractionAscentPermit       : BOOL;

    // === Usage effectif d'un override/bypass de POSITION (consommé PRG_03 → FB_Modes) ===
    // Producteur unique : PRG_04_Treuils_Benne §5. Lecteur : PRG_03_Modes_Cycle (lag 1 scan assumé,
    // même doctrine que les autres échanges PRG_03/PRG_04 de ce bus).
    // TRUE = la limite de position de cet axe est actuellement levée au-delà du nominal :
    // override FDC logiciel N1 maintenu OU bypass N2 effectif de la famille position
    // (TopLimitSwitch / TopLimitSoftware / CableLimitSwitch / LimitLegal / MecaD).
    // Sert à armer le re-homing obligatoire (AF-05 §4bis) — n'est PAS un permis de mouvement.
    PositionLimitOverriddenM1    : BOOL;               // 🧭 Treuil M1 — limite de position levée
    PositionLimitOverriddenM2    : BOOL;               // 🧭 Treuil M2 — limite de position levée

    // === 🕵️ Trace de blocage terrain (consommée FB_TroubleshootingView) ===
    TraceM1                      : ST_TraceWinch;      // 🕵️ Trace blocage treuil M1 (cause priorisée + horodatage)
    TraceM2                      : ST_TraceWinch;      // 🕵️ Trace blocage treuil M2 (cause priorisée + horodatage)

    // === 🔗 ATOMICITÉ BOTH : diagnostic IHM lecture seule ===
    // Permis agrégés consommés par la commande both + cause priorisée du blocage.
    // Aucune action de conduite n'en dépend (l'arrêt est porté par §5/§6 de PRG_04).
    BothActive                   : BOOL;               // 🔗 Intention both active (M1+M2 ensemble)
    BothBlocked                  : BOOL;               // 🔗 Commande Both bloquée par le permis agrégé (diagnostic uniquement)
    BothBlockReason              : E_WinchTraceBlockReason; // 🔗 Cause priorisée du blocage Both

    // === 🚦 Disponibilité de mouvement par axe/sens (base honnête de ArmingPermit) ===
    // Producteur unique : PRG_04_Treuils_Benne §5-0. Lecteurs : PRG_02 (ArmingPermit),
    // FB_TroubleshootingView / IHM (diagnostic « pourquoi ça n'arme pas »).
    ArmingAvailability           : ST_ArmingAvailability;
END_STRUCT
END_TYPE

(* ---- ST_WinchState.st ---- *)
(* ═══════════════════════════════════════════════════════════════
   🚦 ST_WinchState — États, mesures et diagnostics HMI pour un Treuil M1/M2
   ───────────────────────────────────────────────────────────────
   🎨 Destiné aux retours d'informations et bargraphes HMI.
   ═══════════════════════════════════════════════════════════════ *)
TYPE ST_WinchState :
STRUCT
    (* 🚦 États & Mesures (Lecture seule) *)
    Position_M              : REAL;             (* 📊 Position actuelle du câble (mètres) *)
    MeasuredSpeed_Mps       : REAL;             (* 📏 Vitesse linéaire mesurée du câble (m/s), valeur absolue *)
    SpeedDelta_Mps          : REAL;             (* 🔍 Variation de vitesse entre deux scans (m/s) *)
    SpeedVariationDetected  : BOOL;             (* 🔍 Seuil de variation dépassé sur le scan courant *)
    SpeedVariationConfirmed : BOOL;             (* 🛡️ Variation confirmée pendant la durée paramétrée *)
    SpeedStable             : BOOL;             (* 🟢 Vitesse stable pendant la durée paramétrée *)
    SpeedMonitorError       : BOOL;             (* Défaut mémorisé du moniteur vitesse *)
    SpeedMonitorErrorId     : WORD;             (* ❌ Bitfield du moniteur vitesse *)
    EstimatedLoadPct        : REAL;             (* 📊 Estimation empirique, non certifiée *)
    LoadEstimateConfigured  : BOOL;             (* 🟢 Table charge validée pour lecture *)
    SpeedGuardLimited       : BOOL;             (* 🛡️ Palier limité par vitesse réelle *)
    SpeedCmd_Pct            : REAL;             (* 📈 Commande de vitesse finale après rampe (%) *)
    StepNumber              : INT;              (* 🔢 Palier de vitesse actif (0..5) *)
    FBState                 : E_State;          (* 🤖 État de l'automate interne (FB_Winch) *)
    AxisBlockReason         : E_WinchTraceBlockReason; (* 🧩 Cause prioritaire de blocage (miroir de TraceMx.BlockReason) *)
    Ready                   : BOOL;             (* 🟢 Treuil prêt à fonctionner *)
    Busy                    : BOOL;             (* ⚙️ Mouvement en cours *)
    Done                    : BOOL;             (* ✅ Action terminée *)
    Error                   : BOOL;             (* Treuil en défaut *)
    ErrorId                 : WORD;             (* ❌ Code bitfield du défaut treuil *)

    (* 🔌 Sorties Physiques / Indicateurs LEDs *)
    RelayFwd                : BOOL;             (* 🛗 Relais Ascending activé *)
    RelayRev                : BOOL;             (* 🛗 Relais Descending activé *)
    Contactor1              : BOOL;             (* 🔌 Contacteur vitesse palier 1 *)
    Contactor2              : BOOL;             (* 🔌 Contacteur vitesse palier 2 *)
    Contactor3              : BOOL;             (* 🔌 Contacteur vitesse palier 3 *)
    Contactor4              : BOOL;             (* 🔌 Contacteur vitesse palier 4 *)
    BrakeCmd                : BOOL;             (* 🔓 Commande frein (TRUE = desserré / libre) *)
    FinalInterlockState     : E_WinchFinalInterlockState; (* 🛡️ État final lecture seule *)
    FinalInterlockReason    : E_WinchFinalInterlockReason; (* 🛡️ Cause finale mémorisée *)
    FinalInterlockError     : BOOL;             (* 🛡️ Défaut final mémorisé *)
    FinalInterlockErrorId   : WORD;             (* 🛡️ Bitfield final *)
    FinalRestartInhibit     : BOOL;             (* 🔒 Reset + neutre + nouvelle demande obligatoires *)
    FinalRestartRequired    : BOOL;             (* 🔒 Purge anti-redemarrage armee : AuthorizedStep force a 0 tant que non purgee (distinct de RestartInhibit) *)
    FinalMotorRequest       : BOOL;             (* 🔒 Demande moteur vue par la barriere finale (palier>0 ET un seul sens) *)
    FinalNeutralRequestSeen : BOOL;             (* 🔒 Passage au neutre observe pendant un RestartInhibit *)
    BrakeCommandOpenConfirmed : BOOL;           (* 🔌 Contacteur/bobine desserrage confirmé, pas frein mécanique *)
    FinalAuthorizedStep     : INT;              (* 🪜 Palier réellement autorisé *)
    FinalBrakeTimeoutElapsed : TIME;            (* ⏱️ Écoulé watchdog 500ms *)
    FinalRestartDelayElapsed : TIME;            (* ⏱️ Écoulé verrou redémarrage 900ms *)
    FinalStepDelayElapsed    : TIME;            (* ⏱️ Écoulé entre paliers 1s250 *)

    (* 🛡️ Sécurités & Diagnostics *)
    Encoder                 : ST_EncoderHMI;    (* 🧲 Données d'échange et diagnostic du codeur — porte aussi les 9 champs Homing* (voir ST_EncoderHMI) *)

    (* 🔍 Diagnostics de cohérence contacteurs réutilisés *)
    ContactorsCheck         : ST_ContactorCheck; (* 🔌 Coherence contacteurs sens+vitesse *)
    BrakeContactorCheck     : ST_ContactorCheck; (* 🔌 Coherence retour frein *)
    InhibitActive           : BOOL;             (* miroir lecture seule — inhibition arbitrée *)

    (* 🐢 : ralentissement sur bordure — diagnostic zone/limite active *)
    BottomLimitActiveM      : REAL;             (* 📏 Limite basse active (m) — câble physique OU légale, la plus restrictive *)
    InTopSlowdownZone       : BOOL;             (* 🐢 Palier plafonné à 1 : approche limite haute *)
    InBottomSlowdownZone    : BOOL;             (* 🐢 Palier plafonné à 1 : approche limite basse (câble ou légale) *)

    (* 🩺 Diagnostic délai ressenti à la remontée *)
    CommandedAscent           : BOOL;          (* 🩺 Sens interne mémorisé FB_Winch : montée *)
    CommandedDescend          : BOOL;          (* 🩺 Sens interne mémorisé FB_Winch : descente *)
    DirectionChangeDelayElapsed : TIME;         (* 🩺 Écoulé de l'interlock changement/reprise de sens *)
    DirectionChangePending      : BOOL;         (* 🩺 TRUE tant que CommandedDirection n'a pas rejoint Direction *)
END_STRUCT
END_TYPE

(* ---- ST_WinchSymmetryHMI.st ---- *)
TYPE ST_WinchSymmetryHMI :
STRUCT
    BtnReset : BOOL;
    SymmetryOk : BOOL;
    SymmetryValid : BOOL;
    DeltaStartDelay_Ms : UDINT;
    DeltaBrakeReleaseTime_Ms : UDINT;
    DeltaBrakeApplyTime_Ms : UDINT;
    DeltaStopDistance_M : REAL;
    DeltaStopTime_Ms : UDINT;
    MaxSyncDeviation_M : REAL;
END_STRUCT
END_TYPE
